// TIA Portal V21 export
// export: Created 2026-11-08T21:35:27.6716818Z, ExportSetting WithDefaults, DisplayName Totally Integrated Automation Portal, DisplayVersion V21 Update 3, DisplayName STEP 7 Professional, DisplayVersion V21 Update 3, DisplayName STEP 7 Safety, DisplayVersion V21, DisplayName Tech WebApplication, DisplayVersion V21, DisplayName WinCC Basic/Comfort/Advanced, DisplayVersion V21 Update 3, DisplayName WinCC Unified, DisplayVersion V21 Update 3
FUNCTION_BLOCK "FB_StlC_025"   // FB50, STL
TITLE = STL call MOVE
{ S7_Optimized_Access := 'TRUE' }
VERSION : 0.1
// stored: AutoNumber true, IsRetainMemResEnabled false, MemoryReserve 100, UDAEnableTagReadback false
   VAR_INPUT
      "a" : Bool;
      i1 : Int;
      i2 : Int;
      di1 : DInt;
      r1 : Real;
      w1 : Word;
      dw1 : DWord;
      b1 : Byte;
      u1 : UInt;
      ud1 : UDInt;
   END_VAR
   VAR_OUTPUT
      q : Bool;
      io : Int;
      dio : DInt;
      ro : Real;
      wo : Word;
      dwo : DWord;
      bo : Byte;
      udo : UDInt;
   END_VAR
   VAR
      src : Array[0..9] of Int;
      dst : Array[0..9] of Int;
      bits : Array[0..31] of Bool;
      bytes : Array[0..9] of Byte;
      err { S7_SetPoint := 'True'} : ErrorStruct;
      rt : LReal;
   END_VAR
BEGIN

NETWORK
TITLE = 025 MOVE
      CALL  MOVE
      ( IN  := #i1,
        OUT := #io
      );
END_FUNCTION_BLOCK
